(* IEC 61131-3 sources: volt/packages/volt-lsp-iec/test-corpus/pro2193/Device/Plc Logic/Application/09 Misc/Library Manager/ElementCollections, 99 files *)

(* ---- COLLECTION_ERROR.dut ---- *)
TYPE COLLECTION_ERROR :
(
	NO_ERROR := 0,
	NO_MORE_ELEMENTS := 2,
	MAXIMUM_SIZE_OF_ELEMENTS_EXCEEDED,
	NULL_POINTER,
	MAXIMUM_ELEMENT_POSITION_EXCEEDED,
	NOT_FOUND,
	UNSUPPORTED_OPERATION,
	KEY_EXISTS,
	ELEMENT_COUNT_NOT_EQUAL_COUNTER,
	LIST_ITERATOR_EXPECTED,
	LINKED_LIST_ITERATOR_EXPECTED,
	COLLECTION_CHANGED,
	NOT_INITIALIZED,
	ELEMENT_IS_REFERENCED,
	ITREE_NODE_EXPECTED,
	FB_CREATE_ERROR,
	ROOT_NODE_CAN_NOT_BE_MOVED,
	INTERNAL_ERROR,
	NODE_CAN_NOT_BE_MOVED_TO_SUBNODE,
	REALLOC_FAILED
);
END_TYPE

(* ---- KEYVALUEPAIR.dut ---- *)
TYPE KEYVALUEPAIR :
STRUCT
	KEYELEMENT : IElement;
	VALUEELEMENT : IElement;
	NEXT : POINTER TO KeyValuePair;
END_STRUCT
END_TYPE

(* ---- CONSTANTS.gvl ---- *)
VAR_GLOBAL
	GC_TREENODEFACTORY : TreeNodeFactory := STRUCT();
	GC_LINKEDOBJECTREFERENCEFACTORY : LinkedObjectReferenceFactory := STRUCT();
END_VAR

(* ---- VARIABLES.gvl ---- *)
VAR_GLOBAL
	G_LOCKWAITTIME : SYSTIME := 300;
	G_NULLELEMENT : NullElement;
END_VAR

(* ---- IBOOLELEMENT.itf ---- *)
INTERFACE IBOOLELEMENT
END_INTERFACE

(* ---- ICOLLECTION.itf ---- *)
INTERFACE ICOLLECTION
END_INTERFACE

METHOD ADDELEMENT : COLLECTION_ERROR
VAR_INPUT
	ITFELEMENT : IElement;
END_VAR
END_METHOD

METHOD CONTAINSELEMENT : COLLECTION_ERROR
VAR_INPUT
	ITFELEMENT : IElement;
END_VAR
VAR_OUTPUT
	XRESULT : BOOL;
END_VAR
END_METHOD

METHOD COUNTELEMENTS : UDINT
END_METHOD

METHOD ELEMENTITERATOR : COLLECTION_ERROR
VAR_INPUT
	ITFITERATOR : IIterator;
END_VAR
END_METHOD

METHOD REMOVEALLELEMENTS : COLLECTION_ERROR
END_METHOD

METHOD REMOVEELEMENT : COLLECTION_ERROR
VAR_INPUT
	ITFELEMENT : IElement;
END_VAR
END_METHOD

(* ---- ICONTAINSVALUE.itf ---- *)
INTERFACE ICONTAINSVALUE
END_INTERFACE

METHOD CONTAINSVALUE : COLLECTION_ERROR
VAR_INPUT
	ITFELEMENT : IElement;
END_VAR
VAR_OUTPUT
	XRESULT : BOOL;
END_VAR
END_METHOD

(* ---- IDINTELEMENT.itf ---- *)
INTERFACE IDINTELEMENT
END_INTERFACE

(* ---- IDOUBLELINKEDLIST.itf ---- *)
INTERFACE IDOUBLELINKEDLIST
END_INTERFACE

METHOD REMOVEFIRSTELEMENT : COLLECTION_ERROR
END_METHOD

METHOD REMOVELASTELEMENT : COLLECTION_ERROR
END_METHOD

(* ---- IELEMENT.itf ---- *)
INTERFACE IELEMENT
END_INTERFACE

METHOD ELEMENTCOMPARETO : INT
VAR_INPUT
	ITFELEMENT : IElement;
END_VAR
END_METHOD

METHOD ELEMENTEQUALS : BOOL
VAR_INPUT
	ITFELEMENT : IElement;
END_VAR
END_METHOD

METHOD ELEMENTHASHCODE : LINT
END_METHOD

(* ---- IINTELEMENT.itf ---- *)
INTERFACE IINTELEMENT
END_INTERFACE

(* ---- IITERATOR.itf ---- *)
INTERFACE IITERATOR
END_INTERFACE

METHOD HASNEXT : BOOL
END_METHOD

METHOD NEXT : COLLECTION_ERROR
VAR_OUTPUT
	ITFELEMENT : IElement;
END_VAR
END_METHOD

(* ---- ILINKEDLISTITERATOR.itf ---- *)
INTERFACE ILINKEDLISTITERATOR
END_INTERFACE

(* ---- ILINKEDOBJECTREFERENCE.itf ---- *)
INTERFACE ILINKEDOBJECTREFERENCE
END_INTERFACE

(* ---- ILINTELEMENT.itf ---- *)
INTERFACE ILINTELEMENT
END_INTERFACE

(* ---- ILIST.itf ---- *)
INTERFACE ILIST
END_INTERFACE

METHOD GETELEMENTAT : COLLECTION_ERROR
VAR_INPUT
	UDIPOSITION : UDINT;
END_VAR
VAR_OUTPUT
	ITFELEMENT : IElement;
END_VAR
END_METHOD

METHOD GETELEMENTPOSITION : COLLECTION_ERROR
VAR_INPUT
	ITFELEMENT : IElement;
END_VAR
VAR_OUTPUT
	UDIPOSITION : UDINT;
END_VAR
END_METHOD

METHOD INSERTELEMENTAT : COLLECTION_ERROR
VAR_INPUT
	UDIPOSITION : UDINT;
	ITFELEMENT : IElement;
END_VAR
END_METHOD

METHOD REMOVEELEMENTAT : COLLECTION_ERROR
VAR_INPUT
	UDIPOSITION : UDINT;
END_VAR
END_METHOD

METHOD SETELEMENTAT : COLLECTION_ERROR
VAR_INPUT
	UDIPOSITION : UDINT;
	ITFELEMENT : IElement;
END_VAR
END_METHOD

(* ---- ILIST2.itf ---- *)
INTERFACE ILIST2
END_INTERFACE

(* ---- ILISTITERATOR.itf ---- *)
INTERFACE ILISTITERATOR
END_INTERFACE

(* ---- IMAP.itf ---- *)
INTERFACE IMAP
END_INTERFACE

METHOD ADDKEYVALUEPAIR : COLLECTION_ERROR
VAR_INPUT
	ITFKEY : IElement;
	ITFVALUE : IElement;
END_VAR
END_METHOD

METHOD CONTAINSKEY : COLLECTION_ERROR
VAR_INPUT
	ITFKEY : IElement;
END_VAR
VAR_OUTPUT
	XRESULT : BOOL;
END_VAR
END_METHOD

METHOD COUNTKEYS : UDINT
END_METHOD

METHOD GETELEMENTBYKEY : COLLECTION_ERROR
VAR_INPUT
	ITFKEY : IElement;
END_VAR
VAR_OUTPUT
	ITFVALUE : IElement;
END_VAR
END_METHOD

METHOD KEYS : COLLECTION_ERROR
VAR_INPUT
	ITFITERATOR : IIterator;
END_VAR
END_METHOD

METHOD REMOVEBYKEY : COLLECTION_ERROR
VAR_INPUT
	ITFKEY : IElement;
END_VAR
END_METHOD

METHOD VALUES : COLLECTION_ERROR
VAR_INPUT
	ITFITERATOR : IIterator;
END_VAR
END_METHOD

(* ---- IMAP2.itf ---- *)
INTERFACE IMAP2
END_INTERFACE

METHOD REMOVEALLELEMENTS : COLLECTION_ERROR
END_METHOD

(* ---- IMODCOUNTER.itf ---- *)
INTERFACE IMODCOUNTER
END_INTERFACE

(* ---- INULLELEMENT.itf ---- *)
INTERFACE INULLELEMENT
END_INTERFACE

(* ---- IOBJECTREFERENCE.itf ---- *)
INTERFACE IOBJECTREFERENCE
END_INTERFACE

(* ---- IONLINECHANGESAFELINKEDLISTELEMENT.itf ---- *)
INTERFACE IONLINECHANGESAFELINKEDLISTELEMENT
END_INTERFACE

METHOD UPDATEELEMENT
VAR_INPUT
	ITFELEMENT : IElement;
END_VAR
END_METHOD

(* ---- IQUEUE.itf ---- *)
INTERFACE IQUEUE
END_INTERFACE

METHOD PEEK : COLLECTION_ERROR
VAR_OUTPUT
	ITFELEMENT : IElement;
END_VAR
END_METHOD

METHOD POLL : COLLECTION_ERROR
VAR_OUTPUT
	ITFELEMENT : IElement;
END_VAR
END_METHOD

(* ---- IQUEUE2.itf ---- *)
INTERFACE IQUEUE2
END_INTERFACE

(* ---- ISORTEDLIST.itf ---- *)
INTERFACE ISORTEDLIST
END_INTERFACE

METHOD ADDELEMENTWITHOUTSORTING : COLLECTION_ERROR
VAR_INPUT
	ITFELEMENT : IElement;
END_VAR
END_METHOD

METHOD SORT : COLLECTION_ERROR
END_METHOD

(* ---- ISORTEDLIST2.itf ---- *)
INTERFACE ISORTEDLIST2
END_INTERFACE

(* ---- ISTACK.itf ---- *)
INTERFACE ISTACK
END_INTERFACE

METHOD PEEK : COLLECTION_ERROR
VAR_OUTPUT
	ITFELEMENT : IElement;
END_VAR
END_METHOD

METHOD POP : COLLECTION_ERROR
VAR_OUTPUT
	ITFELEMENT : IElement;
END_VAR
END_METHOD

(* ---- ISTACK2.itf ---- *)
INTERFACE ISTACK2
END_INTERFACE

(* ---- ISTRINGELEMENT.itf ---- *)
INTERFACE ISTRINGELEMENT
END_INTERFACE

(* ---- ITIMEELEMENT.itf ---- *)
INTERFACE ITIMEELEMENT
END_INTERFACE

(* ---- ITREENODE.itf ---- *)
INTERFACE ITREENODE
END_INTERFACE

METHOD ADDCHILD : COLLECTION_ERROR
VAR_INPUT
	ITFELEMENT : IElement;
END_VAR
VAR_OUTPUT
	ITFTREENODE : ITreeNode;
END_VAR
END_METHOD

METHOD CHILDREN : COLLECTION_ERROR
VAR_INPUT
	ITFITERATOR : IIterator;
END_VAR
END_METHOD

METHOD CONTAINSCHILD : COLLECTION_ERROR
VAR_INPUT
	ITFELEMENT : IElement;
END_VAR
VAR_OUTPUT
	XRESULT : BOOL;
END_VAR
END_METHOD

METHOD COUNTCHILDREN : UDINT
END_METHOD

METHOD MOVENODE : COLLECTION_ERROR
VAR_INPUT
	ITFTARGETTREENODE : ITreeNode;
END_VAR
END_METHOD

METHOD PARENT : COLLECTION_ERROR
VAR_OUTPUT
	ITFPARENT : ITreeNode;
END_VAR
END_METHOD

METHOD REMOVECHILD : COLLECTION_ERROR
VAR_INPUT
	ITFELEMENT : IElement;
END_VAR
END_METHOD

METHOD ROOTNODE : COLLECTION_ERROR
VAR_OUTPUT
	ITFROOTNODE : ITreeNode;
END_VAR
END_METHOD

(* ---- IUDINTELEMENT.itf ---- *)
INTERFACE IUDINTELEMENT
END_INTERFACE

(* ---- IUINTELEMENT.itf ---- *)
INTERFACE IUINTELEMENT
END_INTERFACE

(* ---- IULINTELEMENT.itf ---- *)
INTERFACE IULINTELEMENT
END_INTERFACE

(* ---- IWSTRINGELEMENT.itf ---- *)
INTERFACE IWSTRINGELEMENT
END_INTERFACE

(* ---- COMPARESTRING.pou ---- *)
FUNCTION COMPARESTRING : INT
VAR_INPUT
	PS1 : POINTER TO STRING;
	PS2 : POINTER TO STRING;
END_VAR
END_FUNCTION

(* ---- COMPAREWSTRING.pou ---- *)
FUNCTION COMPAREWSTRING : INT
VAR_INPUT
	PW1 : POINTER TO WSTRING;
	PW2 : POINTER TO WSTRING;
END_VAR
END_FUNCTION

(* ---- GETLIBVERSION.pou ---- *)
FUNCTION GETLIBVERSION : VERSION
END_FUNCTION

(* ---- GETLIBVERSIONNUMBER.pou ---- *)
FUNCTION GETLIBVERSIONNUMBER : DWORD
END_FUNCTION

(* ---- HASHCODEFROMSTRING.pou ---- *)
FUNCTION HASHCODEFROMSTRING : UDINT
VAR_INPUT
	PSIN : POINTER TO STRING;
END_VAR
END_FUNCTION

(* ---- HASHCODEFROMWSTRING.pou ---- *)
FUNCTION HASHCODEFROMWSTRING : UDINT
VAR_INPUT
	PWIN : POINTER TO WSTRING;
END_VAR
END_FUNCTION

(* ---- ISLIBRELEASED.pou ---- *)
FUNCTION ISLIBRELEASED : BOOL
END_FUNCTION

(* ---- BOOLDATA.pou ---- *)
FUNCTION_BLOCK BOOLDATA EXTENDS InstanceData
VAR_INPUT
	XVALUE : BOOL;
END_VAR
END_FUNCTION_BLOCK

(* ---- BOOLELEMENT.pou ---- *)
FUNCTION_BLOCK BOOLELEMENT EXTENDS InstanceBase
VAR_INPUT
	XVALUE : BOOL;
END_VAR
VAR
	BOOLVALUE : BOOL;
END_VAR
END_FUNCTION_BLOCK

METHOD ELEMENTCOMPARETO : INT
VAR_INPUT
	ITFELEMENT : IElement;
END_VAR
END_METHOD

METHOD ELEMENTEQUALS : BOOL
VAR_INPUT
	ITFELEMENT : IElement;
END_VAR
END_METHOD

METHOD ELEMENTHASHCODE : LINT
END_METHOD

METHOD PRVINSTINIT : FBF.ERROR
VAR_INPUT
	ITFDATA : FBF.IData;
END_VAR
END_METHOD

(* ---- BOOLELEMENTFACTORY.pou ---- *)
FUNCTION_BLOCK BOOLELEMENTFACTORY EXTENDS FactoryBase
VAR
	PRVINSTCOUNT : CAA.COUNT;
	PRVINSTPOOLEXTENDSFACTOR : USINT;
	PRVINSTSIZE : CAA.SIZE;
END_VAR
END_FUNCTION_BLOCK

METHOD CREATE : IBoolElement
VAR_INPUT
	XVALUE : BOOL;
END_VAR
VAR_OUTPUT
	EERROR : FBF.ERROR;
END_VAR
END_METHOD

(* ---- DINTDATA.pou ---- *)
FUNCTION_BLOCK DINTDATA EXTENDS InstanceData
VAR_INPUT
	DIVALUE : DINT;
END_VAR
END_FUNCTION_BLOCK

(* ---- DINTELEMENT.pou ---- *)
FUNCTION_BLOCK DINTELEMENT EXTENDS InstanceBase
VAR_INPUT
	DIVALUE : DINT;
END_VAR
VAR
	DINTVALUE : DINT;
END_VAR
END_FUNCTION_BLOCK

METHOD ELEMENTCOMPARETO : INT
VAR_INPUT
	ITFELEMENT : IElement;
END_VAR
END_METHOD

METHOD ELEMENTEQUALS : BOOL
VAR_INPUT
	ITFELEMENT : IElement;
END_VAR
END_METHOD

METHOD ELEMENTHASHCODE : LINT
END_METHOD

METHOD PRVINSTINIT : FBF.ERROR
VAR_INPUT
	ITFDATA : FBF.IData;
END_VAR
END_METHOD

(* ---- DINTELEMENTFACTORY.pou ---- *)
FUNCTION_BLOCK DINTELEMENTFACTORY EXTENDS FactoryBase
VAR
	PRVINSTCOUNT : CAA.COUNT;
	PRVINSTPOOLEXTENDSFACTOR : USINT;
	PRVINSTSIZE : CAA.SIZE;
END_VAR
END_FUNCTION_BLOCK

METHOD CREATE : IDintElement
VAR_INPUT
	DIVALUE : DINT;
END_VAR
VAR_OUTPUT
	EERROR : FBF.ERROR;
END_VAR
END_METHOD

(* ---- HASHTABLE.pou ---- *)
FUNCTION_BLOCK HASHTABLE EXTENDS InstanceBase
VAR_INPUT
	PAELEMENTS : POINTER TO KeyValuePair;
	PALINKEDELEMENTS : POINTER TO KeyValuePair;
	PAITERATORELEMENTS : POINTER TO IElement;
	UDIMAXELEMENTS : UDINT;
END_VAR
VAR
	_UDICOUNT : UDINT;
	_XWPOINTERTOTHIS : __XWORD := THIS;
	_BYLOCK : BYTE;
	_ULINTCOUNTMODS : ULINT;
	_UIGROWFACTOR : UINT := 1;
	_UIPREALLOCATION : UINT := 100;
	COUNTMODIFICATIONS : ULINT;
END_VAR
END_FUNCTION_BLOCK

METHOD ADDKEYVALUEPAIR : COLLECTION_ERROR
VAR_INPUT
	ITFKEY : IElement;
	ITFVALUE : IElement;
END_VAR
END_METHOD

METHOD ADDKEYVALUEPAIRINTERNAL : COLLECTION_ERROR
VAR_INPUT
	ITFKEY : IElement;
	ITFVALUE : IElement;
	XINCREF : BOOL;
END_VAR
END_METHOD

METHOD CONTAINSKEY : COLLECTION_ERROR
VAR_INPUT
	ITFKEY : IElement;
END_VAR
VAR_OUTPUT
	XRESULT : BOOL;
END_VAR
END_METHOD

METHOD CONTAINSKEYINTERNAL : COLLECTION_ERROR
VAR_INPUT
	ITFKEY : IElement;
END_VAR
VAR_OUTPUT
	XRESULT : BOOL;
END_VAR
END_METHOD

METHOD COUNTKEYS : UDINT
END_METHOD

METHOD DISPOSE : BOOL
END_METHOD

METHOD ELEMENTCOMPARETO : INT
VAR_INPUT
	ITFELEMENT : IElement;
END_VAR
END_METHOD

METHOD ELEMENTEQUALS : BOOL
VAR_INPUT
	ITFELEMENT : IElement;
END_VAR
END_METHOD

METHOD ELEMENTHASHCODE : LINT
END_METHOD

METHOD GETARRAYINDEX : UDINT
VAR_INPUT
	ITFKEY : IElement;
END_VAR
END_METHOD

METHOD GETELEMENTBYKEY : COLLECTION_ERROR
VAR_INPUT
	ITFKEY : IElement;
END_VAR
VAR_OUTPUT
	ITFVALUE : IElement;
END_VAR
END_METHOD

METHOD KEYS : COLLECTION_ERROR
VAR_INPUT
	ITFITERATOR : IIterator;
END_VAR
END_METHOD

METHOD LOCK : BOOL
END_METHOD

METHOD NEXTFREELINKEDELEMENT : COLLECTION_ERROR
VAR_OUTPUT
	PKEYVALUEPAIR : POINTER TO KeyValuePair;
END_VAR
END_METHOD

METHOD REALLOC : BOOL
END_METHOD

METHOD RELEASELOCK
END_METHOD

METHOD REMOVEALLELEMENTS : COLLECTION_ERROR
END_METHOD

METHOD REMOVEBYKEY : COLLECTION_ERROR
VAR_INPUT
	ITFKEY : IElement;
END_VAR
END_METHOD

METHOD VALUES : COLLECTION_ERROR
VAR_INPUT
	ITFITERATOR : IIterator;
END_VAR
END_METHOD

METHOD PRVINSTINIT : FBF.ERROR
VAR_INPUT
	ITFDATA : FBF.IData;
END_VAR
END_METHOD

(* ---- HASHTABLEARGS.pou ---- *)
FUNCTION_BLOCK HASHTABLEARGS EXTENDS InstanceData
VAR_INPUT
	PAELEMENTS : POINTER TO KeyValuePair;
	PALINKEDELEMENTS : POINTER TO KeyValuePair;
	PAITERATORELEMENTS : POINTER TO IElement;
	UDIMAXELEMENTS : UDINT;
	UIGROWFACTOR : UINT;
	UIPREALLOCATION : UINT;
END_VAR
END_FUNCTION_BLOCK

(* ---- HASHTABLEFACTORY.pou ---- *)
FUNCTION_BLOCK HASHTABLEFACTORY EXTENDS FactoryBase
VAR
	PRVINSTCOUNT : CAA.COUNT;
	PRVINSTPOOLEXTENDSFACTOR : USINT;
	PRVINSTSIZE : CAA.SIZE;
END_VAR
END_FUNCTION_BLOCK

METHOD CREATE : IMap2
VAR_INPUT
	UDIMAXELEMENTS : UDINT;
END_VAR
VAR_OUTPUT
	EERROR : FBF.ERROR;
END_VAR
END_METHOD

METHOD CREATEDYNAMICHASHTABLE : IMap2
VAR_INPUT
	UDIINITIALSIZE : UDINT;
	UIGROWFACTOR : UINT;
END_VAR
VAR_OUTPUT
	EERROR : FBF.ERROR;
END_VAR
END_METHOD

METHOD CREATEDYNAMICHASHTABLEPREALLOC : IMap2
VAR_INPUT
	UDIINITIALSIZE : UDINT;
	UIGROWFACTOR : UINT;
	UIPREALLOCATION : UINT;
END_VAR
VAR_OUTPUT
	EERROR : FBF.ERROR;
END_VAR
END_METHOD

(* ---- INTDATA.pou ---- *)
FUNCTION_BLOCK INTDATA EXTENDS InstanceData
VAR_INPUT
	IVALUE : INT;
END_VAR
END_FUNCTION_BLOCK

(* ---- INTELEMENT.pou ---- *)
FUNCTION_BLOCK INTELEMENT EXTENDS InstanceBase
VAR_INPUT
	IVALUE : INT;
END_VAR
VAR
	INTVALUE : INT;
END_VAR
END_FUNCTION_BLOCK

METHOD ELEMENTCOMPARETO : INT
VAR_INPUT
	ITFELEMENT : IElement;
END_VAR
END_METHOD

METHOD ELEMENTEQUALS : BOOL
VAR_INPUT
	ITFELEMENT : IElement;
END_VAR
END_METHOD

METHOD ELEMENTHASHCODE : LINT
END_METHOD

METHOD PRVINSTINIT : FBF.ERROR
VAR_INPUT
	ITFDATA : FBF.IData;
END_VAR
END_METHOD

(* ---- INTELEMENTFACTORY.pou ---- *)
FUNCTION_BLOCK INTELEMENTFACTORY EXTENDS FactoryBase
VAR
	PRVINSTCOUNT : CAA.COUNT;
	PRVINSTPOOLEXTENDSFACTOR : USINT;
	PRVINSTSIZE : CAA.SIZE;
END_VAR
END_FUNCTION_BLOCK

METHOD CREATE : IIntElement
VAR_INPUT
	IVALUE : INT;
END_VAR
VAR_OUTPUT
	EERROR : FBF.ERROR;
END_VAR
END_METHOD

(* ---- LINKEDLIST.pou ---- *)
FUNCTION_BLOCK LINKEDLIST EXTENDS InstanceBase
VAR
	_SNAME : STRING := 'LinkedList';
	_RESULT : RTS_IEC_RESULT;
	_XWPOINTERTOTHIS : __XWORD := THIS;
	_BYLOCK : BYTE;
	_ULINTCOUNTMODS : ULINT;
	_ITFFIRSTLINKEDOBJECTREFERENCE : ILinkedObjectReference := 0;
	_ITFLASTLINKEDOBJECTREFERENCE : ILinkedObjectReference := 0;
	_UDICOUNT : UDINT;
	COUNTMODIFICATIONS : ULINT;
END_VAR
END_FUNCTION_BLOCK

METHOD ADDELEMENT : COLLECTION_ERROR
VAR_INPUT
	ITFELEMENT : IElement;
END_VAR
END_METHOD

METHOD ADDELEMENTINTERNAL : COLLECTION_ERROR
VAR_INPUT
	ITFELEMENT : IElement;
	XINCREMENTREFERENCECOUNTER : BOOL;
END_VAR
END_METHOD

METHOD CONTAINSELEMENT : COLLECTION_ERROR
VAR_INPUT
	ITFELEMENT : IElement;
END_VAR
VAR_OUTPUT
	XRESULT : BOOL;
END_VAR
END_METHOD

METHOD COUNTELEMENTS : UDINT
END_METHOD

METHOD DISPOSE : BOOL
END_METHOD

METHOD ELEMENTCOMPARETO : INT
VAR_INPUT
	ITFELEMENT : IElement;
END_VAR
END_METHOD

METHOD ELEMENTEQUALS : BOOL
VAR_INPUT
	ITFELEMENT : IElement;
END_VAR
END_METHOD

METHOD ELEMENTHASHCODE : LINT
END_METHOD

METHOD ELEMENTITERATOR : COLLECTION_ERROR
VAR_INPUT
	ITFITERATOR : IIterator;
END_VAR
END_METHOD

METHOD LOCK : BOOL
END_METHOD

METHOD RELEASELOCK
END_METHOD

METHOD REMOVEALLELEMENTS : COLLECTION_ERROR
END_METHOD

METHOD REMOVEELEMENT : COLLECTION_ERROR
VAR_INPUT
	ITFELEMENT : IElement;
END_VAR
END_METHOD

METHOD REMOVEELEMENTINTERNAL : COLLECTION_ERROR
VAR_INPUT
	ITFELEMENT : IElement;
	XDECREMENTREFERENCECOUNTER : BOOL;
END_VAR
END_METHOD

METHOD REMOVEFIRSTELEMENT : COLLECTION_ERROR
END_METHOD

METHOD REMOVELASTELEMENT : COLLECTION_ERROR
END_METHOD

METHOD PRVINSTINIT : FBF.ERROR
VAR_INPUT
	ITFDATA : FBF.IData;
END_VAR
END_METHOD

(* ---- LINKEDLISTARGS.pou ---- *)
FUNCTION_BLOCK LINKEDLISTARGS EXTENDS InstanceData
END_FUNCTION_BLOCK

(* ---- LINKEDLISTELEMENTBASE.pou ---- *)
FUNCTION_BLOCK LINKEDLISTELEMENTBASE EXTENDS InstanceBase
VAR
	_ITFOBJECTREFERENCE : IObjectReference;
	OBJECTREFERENCE : IObjectReference;
END_VAR
END_FUNCTION_BLOCK

METHOD ELEMENTCOMPARETO : INT
VAR_INPUT
	ITFELEMENT : IElement;
END_VAR
END_METHOD

METHOD ELEMENTEQUALS : BOOL
VAR_INPUT
	ITFELEMENT : IElement;
END_VAR
END_METHOD

METHOD ELEMENTHASHCODE : LINT
END_METHOD

METHOD UPDATEELEMENT
VAR_INPUT
	ITFELEMENT : IElement;
END_VAR
END_METHOD

(* ---- LINKEDLISTFACTORY.pou ---- *)
FUNCTION_BLOCK LINKEDLISTFACTORY EXTENDS FactoryBase
VAR
	PRVINSTCOUNT : CAA.COUNT;
	PRVINSTPOOLEXTENDSFACTOR : USINT;
	PRVINSTSIZE : CAA.SIZE;
END_VAR
END_FUNCTION_BLOCK

METHOD CREATE : IDoubleLinkedList
VAR_OUTPUT
	EERROR : FBF.ERROR;
END_VAR
END_METHOD

(* ---- LINKEDLISTITERATOR.pou ---- *)
FUNCTION_BLOCK LINKEDLISTITERATOR
VAR
	_ITFLINKEDLISTITERATOR : ILinkedObjectReference;
	_MODCOUNTER : IModCounter;
	_ULINTSTARTMODCOUNT : ULINT;
	_XINVALIDDATA : BOOL;
	FIRSTOBJECTREFERENCE : ILinkedObjectReference;
	MODCOUNTER : IModCounter;
END_VAR
END_FUNCTION_BLOCK

METHOD HASNEXT : BOOL
END_METHOD

METHOD NEXT : COLLECTION_ERROR
VAR_OUTPUT
	ITFELEMENT : IElement;
END_VAR
END_METHOD

(* ---- LINKEDOBJECTREFERENCE.pou ---- *)
FUNCTION_BLOCK LINKEDOBJECTREFERENCE EXTENDS InstanceBase
VAR
	_ITFELEMENT : IElement;
	_ITFLASTLINKEDOBJECTREFERENCE : ILinkedObjectReference;
	_ITFNEXTLINKEDOBJECTREFERENCE : ILinkedObjectReference;
	ELEMENT : IElement;
	LAST : ILinkedObjectReference;
	NEXT : ILinkedObjectReference;
END_VAR
END_FUNCTION_BLOCK

METHOD PRVINSTINIT : FBF.ERROR
VAR_INPUT
	ITFDATA : FBF.IData;
END_VAR
END_METHOD

(* ---- LINKEDOBJECTREFERENCEARGS.pou ---- *)
FUNCTION_BLOCK LINKEDOBJECTREFERENCEARGS EXTENDS InstanceData
END_FUNCTION_BLOCK

(* ---- LINKEDOBJECTREFERENCEFACTORY.pou ---- *)
FUNCTION_BLOCK LINKEDOBJECTREFERENCEFACTORY EXTENDS FactoryBase
VAR
	PRVINSTCOUNT : CAA.COUNT;
	PRVINSTPOOLEXTENDSFACTOR : USINT;
	PRVINSTSIZE : CAA.SIZE;
END_VAR
END_FUNCTION_BLOCK

METHOD CREATE : ILinkedObjectReference
VAR_OUTPUT
	EERROR : FBF.ERROR;
END_VAR
END_METHOD

(* ---- LINTDATA.pou ---- *)
FUNCTION_BLOCK LINTDATA EXTENDS InstanceData
VAR_INPUT
	LIVALUE : LINT;
END_VAR
END_FUNCTION_BLOCK

(* ---- LINTELEMENT.pou ---- *)
FUNCTION_BLOCK LINTELEMENT EXTENDS InstanceBase
VAR_INPUT
	LIVALUE : LINT;
END_VAR
VAR
	LINTVALUE : LINT;
END_VAR
END_FUNCTION_BLOCK

METHOD ELEMENTCOMPARETO : INT
VAR_INPUT
	ITFELEMENT : IElement;
END_VAR
END_METHOD

METHOD ELEMENTEQUALS : BOOL
VAR_INPUT
	ITFELEMENT : IElement;
END_VAR
END_METHOD

METHOD ELEMENTHASHCODE : LINT
END_METHOD

METHOD PRVINSTINIT : FBF.ERROR
VAR_INPUT
	ITFDATA : FBF.IData;
END_VAR
END_METHOD

(* ---- LINTELEMENTFACTORY.pou ---- *)
FUNCTION_BLOCK LINTELEMENTFACTORY EXTENDS FactoryBase
VAR
	PRVINSTCOUNT : CAA.COUNT;
	PRVINSTPOOLEXTENDSFACTOR : USINT;
	PRVINSTSIZE : CAA.SIZE;
END_VAR
END_FUNCTION_BLOCK

METHOD CREATE : ILintElement
VAR_INPUT
	LIVALUE : LINT;
END_VAR
VAR_OUTPUT
	EERROR : FBF.ERROR;
END_VAR
END_METHOD

(* ---- LIST.pou ---- *)
FUNCTION_BLOCK LIST EXTENDS InstanceBase
VAR_INPUT
	PAELEMENTS : POINTER TO IElement;
	UDIMAXELEMENTS : UDINT;
END_VAR
VAR
	_DIMAXPOSITION : DINT := -1;
	_SNAME : STRING := 'List';
	RESULT : RTS_IEC_RESULT;
	_XWPOINTERTOTHIS : __XWORD := THIS;
	_BYLOCK : BYTE;
	_ULINTCOUNTMODS : ULINT;
	_UIGROWFACTOR : UINT := 1;
	COUNTMODIFICATIONS : ULINT;
END_VAR
END_FUNCTION_BLOCK

METHOD ADDELEMENT : COLLECTION_ERROR
VAR_INPUT
	ITFELEMENT : IElement;
END_VAR
END_METHOD

METHOD CONTAINSELEMENT : COLLECTION_ERROR
VAR_INPUT
	ITFELEMENT : IElement;
END_VAR
VAR_OUTPUT
	XRESULT : BOOL;
END_VAR
END_METHOD

METHOD CONTAINSVALUE : COLLECTION_ERROR
VAR_INPUT
	ITFELEMENT : IElement;
END_VAR
VAR_OUTPUT
	XRESULT : BOOL;
END_VAR
END_METHOD

METHOD COUNTELEMENTS : UDINT
END_METHOD

METHOD DISPOSE : BOOL
END_METHOD

METHOD ELEMENTCOMPARETO : INT
VAR_INPUT
	ITFELEMENT : IElement;
END_VAR
END_METHOD

METHOD ELEMENTEQUALS : BOOL
VAR_INPUT
	ITFELEMENT : IElement;
END_VAR
END_METHOD

METHOD ELEMENTHASHCODE : LINT
END_METHOD

METHOD ELEMENTITERATOR : COLLECTION_ERROR
VAR_INPUT
	ITFITERATOR : IIterator;
END_VAR
END_METHOD

METHOD GETELEMENTAT : COLLECTION_ERROR
VAR_INPUT
	UDIPOSITION : UDINT;
END_VAR
VAR_OUTPUT
	ITFELEMENT : IElement;
END_VAR
END_METHOD

METHOD GETELEMENTPOSITION : COLLECTION_ERROR
VAR_INPUT
	ITFELEMENT : IElement;
END_VAR
VAR_OUTPUT
	UDIPOSITION : UDINT;
END_VAR
END_METHOD

METHOD INSERTELEMENTAT : COLLECTION_ERROR
VAR_INPUT
	UDIPOSITION : UDINT;
	ITFELEMENT : IElement;
END_VAR
END_METHOD

METHOD LOCK : BOOL
END_METHOD

METHOD REALLOC : BOOL
END_METHOD

METHOD RELEASELOCK
END_METHOD

METHOD REMOVEALLELEMENTS : COLLECTION_ERROR
END_METHOD

METHOD REMOVEALLELEMENTSINTERNAL : COLLECTION_ERROR
END_METHOD

METHOD REMOVEELEMENT : COLLECTION_ERROR
VAR_INPUT
	ITFELEMENT : IElement;
END_VAR
END_METHOD

METHOD REMOVEELEMENTAT : COLLECTION_ERROR
VAR_INPUT
	UDIPOSITION : UDINT;
END_VAR
END_METHOD

METHOD REMOVEELEMENTATINTERNAL : COLLECTION_ERROR
VAR_INPUT
	UDIPOSITION : UDINT;
END_VAR
END_METHOD

METHOD SETELEMENTAT : COLLECTION_ERROR
VAR_INPUT
	UDIPOSITION : UDINT;
	ITFELEMENT : IElement;
END_VAR
END_METHOD

METHOD PRVINSTINIT : FBF.ERROR
VAR_INPUT
	ITFDATA : FBF.IData;
END_VAR
END_METHOD

(* ---- LISTARGS.pou ---- *)
FUNCTION_BLOCK LISTARGS EXTENDS InstanceData
VAR_INPUT
	PAELEMENTS : POINTER TO IElement;
	UDIMAXELEMENTS : UDINT;
	UIGROWFACTOR : UINT;
END_VAR
END_FUNCTION_BLOCK

(* ---- LISTFACTORY.pou ---- *)
FUNCTION_BLOCK LISTFACTORY EXTENDS FactoryBase
VAR
	PRVINSTCOUNT : CAA.COUNT;
	PRVINSTPOOLEXTENDSFACTOR : USINT;
	PRVINSTSIZE : CAA.SIZE;
END_VAR
END_FUNCTION_BLOCK

METHOD CREATE : IList2
VAR_INPUT
	UDIMAXELEMENTS : UDINT;
END_VAR
VAR_OUTPUT
	EERROR : FBF.ERROR;
END_VAR
END_METHOD

METHOD CREATEDYNAMICLIST : IList2
VAR_INPUT
	UDIINITIALSIZE : UDINT;
	UIGROWFACTOR : UINT;
END_VAR
VAR_OUTPUT
	EERROR : FBF.ERROR;
END_VAR
END_METHOD

(* ---- LISTITERATOR.pou ---- *)
FUNCTION_BLOCK LISTITERATOR
VAR
	_DICOUNT : DINT := -1;
	_PAELEMENTS : POINTER TO IElement := 0;
	_DISIZE : DINT;
	_MODCOUNTER : IModCounter;
	_ULINTSTARTMODCOUNT : ULINT;
	ELEMENTARRAY : POINTER TO IElement;
	ELEMENTARRAYSIZE : DINT;
	MODCOUNTER : IModCounter;
END_VAR
END_FUNCTION_BLOCK

METHOD HASNEXT : BOOL
END_METHOD

METHOD NEXT : COLLECTION_ERROR
VAR_OUTPUT
	ITFELEMENT : IElement;
END_VAR
END_METHOD

(* ---- NULLELEMENT.pou ---- *)
FUNCTION_BLOCK NULLELEMENT
END_FUNCTION_BLOCK

METHOD ELEMENTCOMPARETO : INT
VAR_INPUT
	ITFELEMENT : IElement;
END_VAR
END_METHOD

METHOD ELEMENTEQUALS : BOOL
VAR_INPUT
	ITFELEMENT : IElement;
END_VAR
END_METHOD

METHOD ELEMENTHASHCODE : LINT
END_METHOD

(* ---- QUEUE.pou ---- *)
FUNCTION_BLOCK QUEUE EXTENDS InstanceBase
VAR_INPUT
	PAELEMENTS : POINTER TO IElement;
	UDIMAXELEMENTS : UDINT;
END_VAR
VAR
	_DIMAXREARPOSITION : DINT := -1;
	_DIMAXFRONTPOSITION : DINT := -1;
	_SNAME : STRING := 'List';
	RESULT : RTS_IEC_RESULT;
	_XWPOINTERTOTHIS : __XWORD := THIS;
	_BYLOCK : BYTE;
	_ULINTCOUNTMODS : ULINT;
	_UIGROWFACTOR : UINT := 1;
	COUNTMODIFICATIONS : ULINT;
END_VAR
END_FUNCTION_BLOCK

METHOD ADDELEMENT : COLLECTION_ERROR
VAR_INPUT
	ITFELEMENT : IElement;
END_VAR
END_METHOD

METHOD CONTAINSELEMENT : COLLECTION_ERROR
VAR_INPUT
	ITFELEMENT : IElement;
END_VAR
VAR_OUTPUT
	XRESULT : BOOL;
END_VAR
END_METHOD

METHOD CONTAINSVALUE : COLLECTION_ERROR
VAR_INPUT
	ITFELEMENT : IElement;
END_VAR
VAR_OUTPUT
	XRESULT : BOOL;
END_VAR
END_METHOD

METHOD COUNTELEMENTS : UDINT
END_METHOD

METHOD DISPOSE : BOOL
END_METHOD

METHOD ELEMENTCOMPARETO : INT
VAR_INPUT
	ITFELEMENT : IElement;
END_VAR
END_METHOD

METHOD ELEMENTEQUALS : BOOL
VAR_INPUT
	ITFELEMENT : IElement;
END_VAR
END_METHOD

METHOD ELEMENTHASHCODE : LINT
END_METHOD

METHOD ELEMENTITERATOR : COLLECTION_ERROR
VAR_INPUT
	ITFITERATOR : IIterator;
END_VAR
END_METHOD

METHOD LOCK : BOOL
END_METHOD

METHOD PEEK : COLLECTION_ERROR
VAR_OUTPUT
	ITFELEMENT : IElement;
END_VAR
END_METHOD

METHOD POLL : COLLECTION_ERROR
VAR_OUTPUT
	ITFELEMENT : IElement;
END_VAR
END_METHOD

METHOD REALLOC : BOOL
END_METHOD

METHOD RELEASELOCK
END_METHOD

METHOD REMOVEALLELEMENTS : COLLECTION_ERROR
END_METHOD

METHOD REMOVEALLELEMENTSINTERNAL : COLLECTION_ERROR
END_METHOD

METHOD REMOVEELEMENT : COLLECTION_ERROR
VAR_INPUT
	ITFELEMENT : IElement;
END_VAR
END_METHOD

METHOD REMOVEELEMENTATINTERNAL : COLLECTION_ERROR
VAR_INPUT
	UDIPOSITION : UDINT;
END_VAR
END_METHOD

METHOD PRVINSTINIT : FBF.ERROR
VAR_INPUT
	ITFDATA : FBF.IData;
END_VAR
END_METHOD

(* ---- QUEUEFACTORY.pou ---- *)
FUNCTION_BLOCK QUEUEFACTORY EXTENDS FactoryBase
VAR
	PRVINSTCOUNT : CAA.COUNT;
	PRVINSTPOOLEXTENDSFACTOR : USINT;
	PRVINSTSIZE : CAA.SIZE;
END_VAR
END_FUNCTION_BLOCK

METHOD CREATE : IQueue2
VAR_INPUT
	UDIMAXELEMENTS : UDINT;
END_VAR
VAR_OUTPUT
	EERROR : FBF.ERROR;
END_VAR
END_METHOD

METHOD CREATEDYNAMICQUEUE : IQueue2
VAR_INPUT
	UDIINITIALSIZE : UDINT;
	UIGROWFACTOR : UINT;
END_VAR
VAR_OUTPUT
	EERROR : FBF.ERROR;
END_VAR
END_METHOD

(* ---- SORTEDLIST.pou ---- *)
FUNCTION_BLOCK SORTEDLIST EXTENDS InstanceBase
VAR_INPUT
	PAELEMENTS : POINTER TO IElement;
	UDIMAXELEMENTS : UDINT;
	XSORTAFTERONLINECHANGE : BOOL := FALSE;
END_VAR
VAR
	_DIMAXPOSITION : DINT := -1;
	_SNAME : STRING := 'List';
	RESULT : RTS_IEC_RESULT;
	_XWPOINTERTOTHIS : __XWORD := THIS;
	_BYLOCK : BYTE;
	_HEVT_ONLINECHANGEDONE : RTS_IEC_HANDLE;
	_HINTERFACEEVT_ONLINECHANGEDONE : RTS_IEC_HANDLE;
	_ITFEVENTCALLBACK : CmpEventMgr_Interfaces.ICmpEventCallback;
	_ULINTCOUNTMODS : ULINT;
	_UIGROWFACTOR : UINT := 1;
	COUNTMODIFICATIONS : ULINT;
END_VAR
END_FUNCTION_BLOCK

METHOD ADDELEMENT : COLLECTION_ERROR
VAR_INPUT
	ITFELEMENT : IElement;
END_VAR
END_METHOD

METHOD ADDELEMENTWITHOUTSORTING : COLLECTION_ERROR
VAR_INPUT
	ITFELEMENT : IElement;
END_VAR
END_METHOD

METHOD CONTAINSELEMENT : COLLECTION_ERROR
VAR_INPUT
	ITFELEMENT : IElement;
END_VAR
VAR_OUTPUT
	XRESULT : BOOL;
END_VAR
END_METHOD

METHOD CONTAINSVALUE : COLLECTION_ERROR
VAR_INPUT
	ITFELEMENT : IElement;
END_VAR
VAR_OUTPUT
	XRESULT : BOOL;
END_VAR
END_METHOD

METHOD COUNTELEMENTS : UDINT
END_METHOD

METHOD DISPOSE : BOOL
END_METHOD

METHOD ELEMENTCOMPARETO : INT
VAR_INPUT
	ITFELEMENT : IElement;
END_VAR
END_METHOD

METHOD ELEMENTEQUALS : BOOL
VAR_INPUT
	ITFELEMENT : IElement;
END_VAR
END_METHOD

METHOD ELEMENTHASHCODE : LINT
END_METHOD

METHOD ELEMENTITERATOR : COLLECTION_ERROR
VAR_INPUT
	ITFITERATOR : IIterator;
END_VAR
END_METHOD

METHOD EVENTCALLBACK : UDINT
VAR_INPUT
	PEVENTPARAM : POINTER TO EventParam;
END_VAR
END_METHOD

METHOD FB_INIT : BOOL
VAR_INPUT
	BINITRETAINS : BOOL;
	BINCOPYCODE : BOOL;
END_VAR
END_METHOD

METHOD FB_EXIT : BOOL
VAR_INPUT
	BINCOPYCODE : BOOL;
END_VAR
END_METHOD

METHOD GETELEMENTAT : COLLECTION_ERROR
VAR_INPUT
	UDIPOSITION : UDINT;
END_VAR
VAR_OUTPUT
	ITFELEMENT : IElement;
END_VAR
END_METHOD

METHOD GETELEMENTPOSITION : COLLECTION_ERROR
VAR_INPUT
	ITFELEMENT : IElement;
END_VAR
VAR_OUTPUT
	UDIPOSITION : UDINT;
END_VAR
END_METHOD

METHOD INSERTELEMENTAT : COLLECTION_ERROR
VAR_INPUT
	UDIPOSITION : UDINT;
	ITFELEMENT : IElement;
END_VAR
END_METHOD

METHOD LOCK : BOOL
END_METHOD

METHOD QSORTHELPER : BOOL
VAR_INPUT
	DILEFT : DINT;
	DIRIGHT : DINT;
END_VAR
END_METHOD

METHOD QUICKSORT : BOOL
VAR_INPUT
	DILEFT : DINT;
	DIRIGHT : DINT;
END_VAR
END_METHOD

METHOD REALLOC : BOOL
END_METHOD

METHOD RELEASELOCK
END_METHOD

METHOD REMOVEALLELEMENTS : COLLECTION_ERROR
END_METHOD

METHOD REMOVEALLELEMENTSINTERNAL : COLLECTION_ERROR
END_METHOD

METHOD REMOVEELEMENT : COLLECTION_ERROR
VAR_INPUT
	ITFELEMENT : IElement;
END_VAR
END_METHOD

METHOD REMOVEELEMENTAT : COLLECTION_ERROR
VAR_INPUT
	UDIPOSITION : UDINT;
END_VAR
END_METHOD

METHOD REMOVEELEMENTATINTERNAL : COLLECTION_ERROR
VAR_INPUT
	UDIPOSITION : UDINT;
END_VAR
END_METHOD

METHOD SETELEMENTAT : COLLECTION_ERROR
VAR_INPUT
	UDIPOSITION : UDINT;
	ITFELEMENT : IElement;
END_VAR
END_METHOD

METHOD SORT : COLLECTION_ERROR
END_METHOD

METHOD PRVINSTINIT : FBF.ERROR
VAR_INPUT
	ITFDATA : FBF.IData;
END_VAR
END_METHOD

(* ---- SORTEDLISTFACTORY.pou ---- *)
FUNCTION_BLOCK SORTEDLISTFACTORY EXTENDS FactoryBase
VAR
	PRVINSTCOUNT : CAA.COUNT;
	PRVINSTPOOLEXTENDSFACTOR : USINT;
	PRVINSTSIZE : CAA.SIZE;
END_VAR
END_FUNCTION_BLOCK

METHOD CREATE : ISortedList2
VAR_INPUT
	UDIMAXELEMENTS : UDINT;
END_VAR
VAR_OUTPUT
	EERROR : FBF.ERROR;
END_VAR
END_METHOD

METHOD CREATEDYNAMICLIST : ISortedList2
VAR_INPUT
	UDIINITIALSIZE : UDINT;
	UIGROWFACTOR : UINT;
END_VAR
VAR_OUTPUT
	EERROR : FBF.ERROR;
END_VAR
END_METHOD

(* ---- STACK.pou ---- *)
FUNCTION_BLOCK STACK EXTENDS InstanceBase
VAR_INPUT
	PAELEMENTS : POINTER TO IElement;
	UDIMAXELEMENTS : UDINT;
END_VAR
VAR
	_DIMAXPOSITION : DINT := -1;
	_SNAME : STRING := 'List';
	RESULT : RTS_IEC_RESULT;
	_XWPOINTERTOTHIS : __XWORD := THIS;
	_BYLOCK : BYTE;
	_ULINTCOUNTMODS : ULINT;
	_UIGROWFACTOR : UINT := 1;
	COUNTMODIFICATIONS : ULINT;
END_VAR
END_FUNCTION_BLOCK

METHOD ADDELEMENT : COLLECTION_ERROR
VAR_INPUT
	ITFELEMENT : IElement;
END_VAR
END_METHOD

METHOD CONTAINSELEMENT : COLLECTION_ERROR
VAR_INPUT
	ITFELEMENT : IElement;
END_VAR
VAR_OUTPUT
	XRESULT : BOOL;
END_VAR
END_METHOD

METHOD CONTAINSVALUE : COLLECTION_ERROR
VAR_INPUT
	ITFELEMENT : IElement;
END_VAR
VAR_OUTPUT
	XRESULT : BOOL;
END_VAR
END_METHOD

METHOD COUNTELEMENTS : UDINT
END_METHOD

METHOD DISPOSE : BOOL
END_METHOD

METHOD ELEMENTCOMPARETO : INT
VAR_INPUT
	ITFELEMENT : IElement;
END_VAR
END_METHOD

METHOD ELEMENTEQUALS : BOOL
VAR_INPUT
	ITFELEMENT : IElement;
END_VAR
END_METHOD

METHOD ELEMENTHASHCODE : LINT
END_METHOD

METHOD ELEMENTITERATOR : COLLECTION_ERROR
VAR_INPUT
	ITFITERATOR : IIterator;
END_VAR
END_METHOD

METHOD LOCK : BOOL
END_METHOD

METHOD PEEK : COLLECTION_ERROR
VAR_OUTPUT
	ITFELEMENT : IElement;
END_VAR
END_METHOD

METHOD POP : COLLECTION_ERROR
VAR_OUTPUT
	ITFELEMENT : IElement;
END_VAR
END_METHOD

METHOD REALLOC : BOOL
END_METHOD

METHOD RELEASELOCK
END_METHOD

METHOD REMOVEALLELEMENTS : COLLECTION_ERROR
END_METHOD

METHOD REMOVEALLELEMENTSINTERNAL : COLLECTION_ERROR
END_METHOD

METHOD REMOVEELEMENT : COLLECTION_ERROR
VAR_INPUT
	ITFELEMENT : IElement;
END_VAR
END_METHOD

METHOD REMOVEELEMENTATINTERNAL : COLLECTION_ERROR
VAR_INPUT
	UDIPOSITION : UDINT;
END_VAR
END_METHOD

METHOD PRVINSTINIT : FBF.ERROR
VAR_INPUT
	ITFDATA : FBF.IData;
END_VAR
END_METHOD

(* ---- STACKFACTORY.pou ---- *)
FUNCTION_BLOCK STACKFACTORY EXTENDS FactoryBase
VAR
	PRVINSTCOUNT : CAA.COUNT;
	PRVINSTPOOLEXTENDSFACTOR : USINT;
	PRVINSTSIZE : CAA.SIZE;
END_VAR
END_FUNCTION_BLOCK

METHOD CREATE : IStack2
VAR_INPUT
	UDIMAXELEMENTS : UDINT;
END_VAR
VAR_OUTPUT
	EERROR : FBF.ERROR;
END_VAR
END_METHOD

METHOD CREATEDYNAMICSTACK : IStack2
VAR_INPUT
	UDIINITIALSIZE : UDINT;
	UIGROWFACTOR : UINT;
END_VAR
VAR_OUTPUT
	EERROR : FBF.ERROR;
END_VAR
END_METHOD

(* ---- STRINGDATA.pou ---- *)
FUNCTION_BLOCK STRINGDATA EXTENDS InstanceData
VAR_INPUT
	SVALUE : STRING;
END_VAR
END_FUNCTION_BLOCK

(* ---- STRINGELEMENT.pou ---- *)
FUNCTION_BLOCK STRINGELEMENT EXTENDS InstanceBase
VAR_INPUT
	SVALUE : STRING;
END_VAR
VAR
	STRINGVALUE : STRING;
END_VAR
END_FUNCTION_BLOCK

METHOD ELEMENTCOMPARETO : INT
VAR_INPUT
	ITFELEMENT : IElement;
END_VAR
END_METHOD

METHOD ELEMENTEQUALS : BOOL
VAR_INPUT
	ITFELEMENT : IElement;
END_VAR
END_METHOD

METHOD ELEMENTHASHCODE : LINT
END_METHOD

METHOD PRVINSTINIT : FBF.ERROR
VAR_INPUT
	ITFDATA : FBF.IData;
END_VAR
END_METHOD

(* ---- STRINGELEMENTFACTORY.pou ---- *)
FUNCTION_BLOCK STRINGELEMENTFACTORY EXTENDS FactoryBase
VAR
	PRVINSTCOUNT : CAA.COUNT;
	PRVINSTPOOLEXTENDSFACTOR : USINT;
	PRVINSTSIZE : CAA.SIZE;
END_VAR
END_FUNCTION_BLOCK

METHOD CREATE : IStringElement
VAR_INPUT
	SVALUE : STRING;
END_VAR
VAR_OUTPUT
	EERROR : FBF.ERROR;
END_VAR
END_METHOD

(* ---- TIMEDATA.pou ---- *)
FUNCTION_BLOCK TIMEDATA EXTENDS InstanceData
VAR_INPUT
	TVALUE : TIME;
END_VAR
END_FUNCTION_BLOCK

(* ---- TIMEELEMENT.pou ---- *)
FUNCTION_BLOCK TIMEELEMENT EXTENDS InstanceBase
VAR_INPUT
	TVALUE : TIME;
END_VAR
VAR
	TIMEVALUE : TIME;
END_VAR
END_FUNCTION_BLOCK

METHOD ELEMENTCOMPARETO : INT
VAR_INPUT
	ITFELEMENT : IElement;
END_VAR
END_METHOD

METHOD ELEMENTEQUALS : BOOL
VAR_INPUT
	ITFELEMENT : IElement;
END_VAR
END_METHOD

METHOD ELEMENTHASHCODE : LINT
END_METHOD

METHOD PRVINSTINIT : FBF.ERROR
VAR_INPUT
	ITFDATA : FBF.IData;
END_VAR
END_METHOD

(* ---- TIMEELEMENTFACTORY.pou ---- *)
FUNCTION_BLOCK TIMEELEMENTFACTORY EXTENDS FactoryBase
VAR
	PRVINSTCOUNT : CAA.COUNT;
	PRVINSTPOOLEXTENDSFACTOR : USINT;
	PRVINSTSIZE : CAA.SIZE;
END_VAR
END_FUNCTION_BLOCK

METHOD CREATE : ITimeElement
VAR_INPUT
	TVALUE : TIME;
END_VAR
VAR_OUTPUT
	EERROR : FBF.ERROR;
END_VAR
END_METHOD

(* ---- TREENODE.pou ---- *)
FUNCTION_BLOCK TREENODE EXTENDS InstanceBase
VAR
	_LINKEDLIST : LinkedList;
	_XWPOINTERTOTHIS : __XWORD := THIS;
	_BYLOCK : BYTE;
	_ITFELEMENT : IElement;
	_ITFPARENTNODE : ITreeNode;
	ELEMENT : IElement;
END_VAR
END_FUNCTION_BLOCK

METHOD ADDCHILD : COLLECTION_ERROR
VAR_INPUT
	ITFELEMENT : IElement;
END_VAR
VAR_OUTPUT
	ITFTREENODE : ITreeNode;
END_VAR
END_METHOD

METHOD CHILDREN : COLLECTION_ERROR
VAR_INPUT
	ITFITERATOR : IIterator;
END_VAR
END_METHOD

METHOD CONTAINSCHILD : COLLECTION_ERROR
VAR_INPUT
	ITFELEMENT : IElement;
END_VAR
VAR_OUTPUT
	XRESULT : BOOL;
END_VAR
END_METHOD

METHOD CONTAINSSUBNODE : COLLECTION_ERROR
VAR_INPUT
	ITFTREENODE : ITreeNode;
END_VAR
VAR_OUTPUT
	XRESULT : BOOL;
END_VAR
END_METHOD

METHOD COUNTCHILDREN : UDINT
END_METHOD

METHOD DISPOSE : BOOL
END_METHOD

METHOD ELEMENTCOMPARETO : INT
VAR_INPUT
	ITFELEMENT : IElement;
END_VAR
END_METHOD

METHOD ELEMENTEQUALS : BOOL
VAR_INPUT
	ITFELEMENT : IElement;
END_VAR
END_METHOD

METHOD ELEMENTHASHCODE : LINT
END_METHOD

METHOD LOCK : BOOL
END_METHOD

METHOD MOVENODE : COLLECTION_ERROR
VAR_INPUT
	ITFTARGETTREENODE : ITreeNode;
END_VAR
END_METHOD

METHOD PARENT : COLLECTION_ERROR
VAR_OUTPUT
	ITFPARENT : ITreeNode;
END_VAR
END_METHOD

METHOD RELEASELOCK
END_METHOD

METHOD REMOVECHILD : COLLECTION_ERROR
VAR_INPUT
	ITFELEMENT : IElement;
END_VAR
END_METHOD

METHOD ROOTNODE : COLLECTION_ERROR
VAR_OUTPUT
	ITFROOTNODE : ITreeNode;
END_VAR
END_METHOD

METHOD PRVINSTINIT : FBF.ERROR
VAR_INPUT
	ITFDATA : FBF.IData;
END_VAR
END_METHOD

(* ---- TREENODEARGS.pou ---- *)
FUNCTION_BLOCK TREENODEARGS EXTENDS InstanceData
VAR_INPUT
	ITFELEMENT : IElement;
	ITFPARENT : ITreeNode;
END_VAR
END_FUNCTION_BLOCK

(* ---- TREENODEFACTORY.pou ---- *)
FUNCTION_BLOCK TREENODEFACTORY EXTENDS FactoryBase
VAR
	PRVINSTCOUNT : CAA.COUNT;
	PRVINSTPOOLEXTENDSFACTOR : USINT;
	PRVINSTSIZE : CAA.SIZE;
END_VAR
END_FUNCTION_BLOCK

METHOD CREATE : ITreeNode
VAR_INPUT
	ITFELEMENT : IElement;
END_VAR
VAR_OUTPUT
	EERROR : FBF.ERROR;
END_VAR
END_METHOD

METHOD CREATEINTERNAL : ITreeNode
VAR_INPUT
	ITFELEMENT : IElement;
	ITFPARENT : ITreeNode;
END_VAR
VAR_OUTPUT
	EERROR : FBF.ERROR;
END_VAR
END_METHOD

(* ---- UDINTDATA.pou ---- *)
FUNCTION_BLOCK UDINTDATA EXTENDS InstanceData
VAR_INPUT
	UDIVALUE : UDINT;
END_VAR
END_FUNCTION_BLOCK

(* ---- UDINTELEMENT.pou ---- *)
FUNCTION_BLOCK UDINTELEMENT EXTENDS InstanceBase
VAR_INPUT
	UDIVALUE : UDINT;
END_VAR
VAR
	UDINTVALUE : UDINT;
END_VAR
END_FUNCTION_BLOCK

METHOD ELEMENTCOMPARETO : INT
VAR_INPUT
	ITFELEMENT : IElement;
END_VAR
END_METHOD

METHOD ELEMENTEQUALS : BOOL
VAR_INPUT
	ITFELEMENT : IElement;
END_VAR
END_METHOD

METHOD ELEMENTHASHCODE : LINT
END_METHOD

METHOD PRVINSTINIT : FBF.ERROR
VAR_INPUT
	ITFDATA : FBF.IData;
END_VAR
END_METHOD

(* ---- UDINTELEMENTFACTORY.pou ---- *)
FUNCTION_BLOCK UDINTELEMENTFACTORY EXTENDS FactoryBase
VAR
	PRVINSTCOUNT : CAA.COUNT;
	PRVINSTPOOLEXTENDSFACTOR : USINT;
	PRVINSTSIZE : CAA.SIZE;
END_VAR
END_FUNCTION_BLOCK

METHOD CREATE : IUdintElement
VAR_INPUT
	UDIVALUE : UDINT;
END_VAR
VAR_OUTPUT
	EERROR : FBF.ERROR;
END_VAR
END_METHOD

(* ---- UINTDATA.pou ---- *)
FUNCTION_BLOCK UINTDATA EXTENDS InstanceData
VAR_INPUT
	UIVALUE : UINT;
END_VAR
END_FUNCTION_BLOCK

(* ---- UINTELEMENT.pou ---- *)
FUNCTION_BLOCK UINTELEMENT EXTENDS InstanceBase
VAR_INPUT
	UIVALUE : UINT;
END_VAR
VAR
	UINTVALUE : UINT;
END_VAR
END_FUNCTION_BLOCK

METHOD ELEMENTCOMPARETO : INT
VAR_INPUT
	ITFELEMENT : IElement;
END_VAR
END_METHOD

METHOD ELEMENTEQUALS : BOOL
VAR_INPUT
	ITFELEMENT : IElement;
END_VAR
END_METHOD

METHOD ELEMENTHASHCODE : LINT
END_METHOD

METHOD PRVINSTINIT : FBF.ERROR
VAR_INPUT
	ITFDATA : FBF.IData;
END_VAR
END_METHOD

(* ---- UINTELEMENTFACTORY.pou ---- *)
FUNCTION_BLOCK UINTELEMENTFACTORY EXTENDS FactoryBase
VAR
	PRVINSTCOUNT : CAA.COUNT;
	PRVINSTPOOLEXTENDSFACTOR : USINT;
	PRVINSTSIZE : CAA.SIZE;
END_VAR
END_FUNCTION_BLOCK

METHOD CREATE : IUintElement
VAR_INPUT
	UIVALUE : UINT;
END_VAR
VAR_OUTPUT
	EERROR : FBF.ERROR;
END_VAR
END_METHOD

(* ---- ULINTDATA.pou ---- *)
FUNCTION_BLOCK ULINTDATA EXTENDS InstanceData
VAR_INPUT
	ULIVALUE : ULINT;
END_VAR
END_FUNCTION_BLOCK

(* ---- ULINTELEMENT.pou ---- *)
FUNCTION_BLOCK ULINTELEMENT EXTENDS InstanceBase
VAR_INPUT
	ULIVALUE : ULINT;
END_VAR
VAR
	ULINTVALUE : ULINT;
END_VAR
END_FUNCTION_BLOCK

METHOD ELEMENTCOMPARETO : INT
VAR_INPUT
	ITFELEMENT : IElement;
END_VAR
END_METHOD

METHOD ELEMENTEQUALS : BOOL
VAR_INPUT
	ITFELEMENT : IElement;
END_VAR
END_METHOD

METHOD ELEMENTHASHCODE : LINT
END_METHOD

METHOD PRVINSTINIT : FBF.ERROR
VAR_INPUT
	ITFDATA : FBF.IData;
END_VAR
END_METHOD

(* ---- ULINTELEMENTFACTORY.pou ---- *)
FUNCTION_BLOCK ULINTELEMENTFACTORY EXTENDS FactoryBase
VAR
	PRVINSTCOUNT : CAA.COUNT;
	PRVINSTPOOLEXTENDSFACTOR : USINT;
	PRVINSTSIZE : CAA.SIZE;
END_VAR
END_FUNCTION_BLOCK

METHOD CREATE : IUlintElement
VAR_INPUT
	ULIVALUE : ULINT;
END_VAR
VAR_OUTPUT
	EERROR : FBF.ERROR;
END_VAR
END_METHOD

(* ---- WSTRINGDATA.pou ---- *)
FUNCTION_BLOCK WSTRINGDATA EXTENDS InstanceData
VAR_INPUT
	WSVALUE : WSTRING;
END_VAR
END_FUNCTION_BLOCK

(* ---- WSTRINGELEMENT.pou ---- *)
FUNCTION_BLOCK WSTRINGELEMENT EXTENDS InstanceBase
VAR_INPUT
	WSVALUE : WSTRING;
END_VAR
VAR
	WSTRINGVALUE : WSTRING;
END_VAR
END_FUNCTION_BLOCK

METHOD ELEMENTCOMPARETO : INT
VAR_INPUT
	ITFELEMENT : IElement;
END_VAR
END_METHOD

METHOD ELEMENTEQUALS : BOOL
VAR_INPUT
	ITFELEMENT : IElement;
END_VAR
END_METHOD

METHOD ELEMENTHASHCODE : LINT
END_METHOD

METHOD PRVINSTINIT : FBF.ERROR
VAR_INPUT
	ITFDATA : FBF.IData;
END_VAR
END_METHOD

(* ---- WSTRINGELEMENTFACTORY.pou ---- *)
FUNCTION_BLOCK WSTRINGELEMENTFACTORY EXTENDS FactoryBase
VAR
	PRVINSTCOUNT : CAA.COUNT;
	PRVINSTPOOLEXTENDSFACTOR : USINT;
	PRVINSTSIZE : CAA.SIZE;
END_VAR
END_FUNCTION_BLOCK

METHOD CREATE : IWStringElement
VAR_INPUT
	WSVALUE : WSTRING;
END_VAR
VAR_OUTPUT
	EERROR : FBF.ERROR;
END_VAR
END_METHOD
